// TIA Portal V21 export
// export: Created 2026-11-10T19:11:33.8315046Z, ExportSetting WithDefaults, DisplayName Totally Integrated Automation Portal, DisplayVersion V21 Update 3, DisplayName STEP 7 Professional, DisplayVersion V21 Update 3, DisplayName STEP 7 Safety, DisplayVersion V21, DisplayName Tech WebApplication, DisplayVersion V21, DisplayName WinCC Basic/Comfort/Advanced, DisplayVersion V21 Update 3, DisplayName WinCC Unified, DisplayVersion V21 Update 3
DATA_BLOCK "DB_TCON"   // DB11
// stored: AutoNumber true, DBAccessibleFromOPCUA true, DBAccessibleFromWebserver true, InstanceOfName TCON, OfSystemLibElement TCON, OfSystemLibVersion 4.0
"TCON"
   // VAR_INPUT
   //    REQ : Bool;
   //    ID : CONN_OUC;
   // END_VAR
   // VAR_OUTPUT
   //    DONE : Bool;
   //    BUSY : Bool;
   //    ERROR : Bool;
   //    STATUS : Word;
   // END_VAR
   // VAR_IN_OUT
   //    CONNECT : Variant;
   // END_VAR
BEGIN
END_DATA_BLOCK
